Fanuc KAREL source: ko00047.KL

-- PROVISIONAL review KL for V770-1; original PC SHA256 167c279da0602ff33929993c5918ff83a4610d81e64dcc48b4d5acb1509dec0b
-- Incomplete behavior may be omitted. Consult companion uncertainty JSON. Do not deploy.
PROGRAM KO00047
%NOLOCKGROUP
BEGIN
  -- UNRESOLVED_PC offsets 5-12; opcodes 9D,23
  -- UNRESOLVED_PC offsets 17-69; opcodes 27,27,49,7E,AD,27,49,7E,AD,22,31,7E,4A
  -- UNRESOLVED_PC offsets 74-78; opcodes 7F
END KO00047
